Fanuc KAREL source: kb00040.compact.KL

PROGRAM KB00040
%STACKSIZE=65535
%PRIORITY=65535
%NOLOCKGROUP
VAR
P1 : STRING[80]
P2 : INTEGER
BEGIN
P1='A'
P2=1
CNV_STR_INT(P1,P2)
END KB00040
